Fanuc KAREL source: ko00077.KL

-- PROVISIONAL review KL for V770-1; original PC SHA256 e9b52fa68e23c49322cd87ff5a9a61454013b0f78c354a6c92741b48397e8033
-- Incomplete behavior may be omitted. Consult companion uncertainty JSON. Do not deploy.
PROGRAM KO00077
%NOLOCKGROUP
BEGIN
  -- UNRESOLVED_PC offsets 5-12; opcodes 9D,23
  -- UNRESOLVED_PC offsets 17-66; opcodes 27,22,1C,27,49,7E,AD,22,31,7E,4A
  -- UNRESOLVED_PC offsets 71-75; opcodes 7F
END KO00077
